// TIA Portal V20 export
// export: Created 2026-10-20T18:55:31.2937871Z, ExportSetting None, DisplayName Totally Integrated Automation Portal, DisplayVersion V20 Update 6, DisplayName TIA Portal Openness, DisplayVersion V20 Update 6, DisplayName TIA Portal Version Control Interface, DisplayVersion V20 Update 6, DisplayName SINAMICS Startdrive Advanced, DisplayVersion V20 SP1, DisplayName SINAMICS Startdrive G130, G150, S120, S150, SINAMICS MV, G220, S200, S210, DisplayVersion V20 SP1, DisplayName SINAMICS Startdrive G110M, G120, G120C, G120D, G120P, G115D, DisplayVersion V20 SP1, DisplayName STEP 7 Professional, DisplayVersion V20 Update 6, DisplayName STEP 7 Safety, DisplayVersion V20 Update 2, DisplayName WinCC Basic/Comfort/Advanced, DisplayVersion V20 Update 6, DisplayName WinCC Unified, DisplayVersion V20 Update 6
VAR_GLOBAL   // PLC tag table "IO_Turck_5"
   "Light_Rear_1_Intensity2(5)" AT %QB1415 : Byte;   // Last byte - 12
   "Light_Rear_1_Color2(5)" AT %QB1417 : Byte;   // Last byte - 10
   "Light_Rear_1_Bounce_Style(5)" AT %QB1413 : Byte;   // Last byte - 14
   "Light_Rear_1_Speed(5)" AT %QB1421 : Byte;   // Last byte - 6
   "Light_Front_1_Percent_Width1(5)" AT %QB1320 : Byte;   // Last byte - 16
   "Light_Front_1_Animation(5)" AT %QB1336 : Byte;   // Last byte
   "Light_Front_1_Speed(5)" AT %QB1330 : Byte;   // Last byte - 6
   "Light_Front_1_Intensity2(5)" AT %QB1324 : Byte;   // Last byte - 12
   "Light_Rear_1_Percent_Width1(5)" AT %QB1411 : Byte;   // Last byte - 16
   "Light_Front_1_1_Direction(5)" AT %QB1318 : Byte;   // Last byte - 18
   "Light_Front_1_Color2(5)" AT %QB1326 : Byte;   // Last byte - 10
   "Light_Rear_1_Color1(5)" AT %QB1425 : Byte;   // Last byte - 2
   "Light_Rear_1_Intensity1(5)" AT %QB1423 : Byte;   // Last byte - 4
   "Light_Rear_1_Animation(5)" AT %QB1427 : Byte;   // Last byte
   "Light_Front_1_Bounce_Style(5)" AT %QB1322 : Byte;   // Last byte - 14
   "Light_Front_1_Color1(5)" AT %QB1334 : Byte;   // Last byte - 2
   "Light_Front_1_Intensity1(5)" AT %QB1332 : Byte;   // Last byte - 4
   "Light_Rear_1_Direction(5)" AT %QB1409 : Byte;   // Last byte - 18
   "Light_Rear_1_Pulse_Pattern(5)" AT %QB1419 : Byte;   // Last byte - 8
   "Light_Front_1_Pulse_Pattern(5)" AT %QB1328 : Byte;   // Last byte - 8
END_VAR
